Staubli VAL3: CalToolPos7.pgx

public program CalToolPos7(tool& x_tTool)
  local frame l_fFrame
  local num l_nFrameErr
  local point l_pCenter
  local bool l_bStatus
  local point l_p5flange
begin
  //定义中心点xyz
  link(l_fFrame,world)
  link(l_pCenter,world)
  //
  call _CalpSphere(db:pTeach1,db:pTeach2,db:pTeach3,db:pTeach4,l_pCenter,l_bStatus)
  l_nFrameErr=setFrame(db:pTeach5,db:pTeach6,db:pTeach7,l_fFrame)
  switch l_nFrameErr
    case 0
      l_pCenter.trsf.rx=l_fFrame.trsf.rx
      l_pCenter.trsf.ry=l_fFrame.trsf.ry
      l_pCenter.trsf.rz=l_fFrame.trsf.rz
      x_tTool.trsf=!db:pTeach5.trsf*l_pCenter.trsf
    break
    case -1,-2
      call db:hmiAlert("DeviationIsTooLarge","warning")
    break
  endSwitch
  call db:hmiAlert("SaveInTool1","info")
end
